(* IEC 61131-3 sources: kns-port-domestic/tools/inventory_tests/fixtures/lib/src/POUs/FB_Base, 3 files *)

(* ---- FB_Base.decl.st ---- *)
// Назначение: абстрактная база с источником времени (SUPER^ и LTIME() в комментарии не считаются)
{attribute 'call_after_init'}
FUNCTION_BLOCK ABSTRACT FB_Base IMPLEMENTS I_Dev
VAR_IN_OUT CONSTANT
    stCfg : ST_Base;
END_VAR
VAR
    ltLast : LTIME;
    itfNext : I_Base;
    refValue : REFERENCE TO DINT;
    pValue : POINTER TO DINT;
    sNote : STRING := 'SUPER^ и __NEW в строке тоже не считаются';
END_VAR
VAR_STAT
    diCount : DINT;
END_VAR

(* ---- FB_Base.impl.st ---- *)
(* LTIME() в блочном комментарии *)
ltLast := LTIME();
pValue := ADR(diCount);
refValue REF= diCount;
IF __ISVALIDREF(refValue) THEN
    diCount := diCount + 1;
END_IF

(* ---- FB_init.method.decl.st ---- *)
METHOD FB_init : BOOL
VAR_INPUT
    bInitRetains : BOOL;
    bInCopyCode : BOOL;
END_VAR
